(*
SPDX-FileCopyrightText: © 2026 Oleksandr Tiutyk <trofimich@gmail.com>
SPDX-License-Identifier: MIT
License: https://opensource.org/license/mit
*)

(*!
<summary>Pairs a path with its expected lexical outcomes for directory and file validation.</summary>
*)
TYPE PATH_VALIDATION_TEST_CASE :
STRUCT
	//! <summary>Null-terminated path passed to each lexical validator.</summary>
	Path : Tc2_System.T_MaxString;
	//! <summary>Expected result from IsValidDirectoryPath.</summary>
	DirectoryAccepted : BOOL;
	//! <summary>Expected result from IsValidFilePath.</summary>
	FileAccepted : BOOL;
END_STRUCT
END_TYPE

(* stored: Version 1.1.0.1
   DUT PATH_VALIDATION_TEST_CASE: Id {480e0279-7f20-47b2-8710-4971d5f17b01} *)
